FUNCTION_BLOCK "FB_ConditionalSelectAndAggregate"
{ S7_Optimized_Access := 'FALSE' }
VERSION : 1.0

VAR_INPUT
    old_z : Int;
END_VAR

VAR_OUTPUT
    newz : Int;
END_VAR

VAR
    ax : Int := 42;
    ay : Int := 333;
END_VAR

BEGIN

    IF NOT (#ax > #old_z) THEN // MUTATED: COND_NEGATE
        #newz := #ay;
    ELSE
        #newz := #old_z;
    END_IF;

    #newz := #newz + #ax + #ay;

END_FUNCTION_BLOCK
